// ============================================================================
// FB_CTD: 减计数器
// 描述: CD上升沿时CV减1, 当CV<=0时Q变为TRUE
// ============================================================================

FUNCTION_BLOCK FB_CTD
VAR_INPUT
    CD   : BOOL;   // 减计数脉冲输入 (上升沿有效)
    LOAD : BOOL;   // 加载预设值 (TRUE时设置CV=PV)
    PV   : INT;    // 预设计数值 (初始加载值)
END_VAR
VAR_OUTPUT
    Q    : BOOL;   // 计数完成输出 (当CV<=0时为TRUE)
    CV   : INT;    // 当前计数值
END_VAR
VAR
    LastCD : BOOL := FALSE;
END_VAR

BEGIN
    // LOAD为TRUE时加载PV到CV
    IF #LOAD THEN
        #CV := #PV;
    ELSIF #CD AND NOT #LastCD THEN
        // CD上升沿且CV>0时减1
        IF #CV > 0 THEN
            #CV := #CV - 1;
        END_IF;
    END_IF;

    // CV<=0时输出TRUE
    #Q := (#CV <= 0);

    // 保存当前CD状态用于下次边沿检测
    #LastCD := #CD;

END_FUNCTION_BLOCK
